(* CODESYS project listofinterface.library
   DefaultNamespace: KOSTAL.TC3.Components.ListOf.Interface
   DocFormat: reStructuredText
   Description: List of Items from base Interface {KOSTAL_TC3_Core_System.I_Interface}
      In addition to the interface, each item contains the pointer to the previous item as well as the pointer to the next item in the list.
   Author: Frank Dümpelmann
   Title: KOSTAL.TC3.Components.ListOf.Interface
   Version: 2019.1.0.0
   Company: KOSTAL GmbH & Co.KG
   Placeholder: KOSTAL.TC3.Components.ListOf.Interface

Project tree, tasks and I/O mapping:
  libraries: KOSTAL.TC3.Core.functionResponse, 2019.0.3.0 (KOSTAL GmbH & Co.KG); KOSTAL.TC3.Core.Settings, 2019.0.1.0 (KOSTAL GmbH & Co.KG); KOSTAL.TC3.Core.System, 2019.0.0.0 (KOSTAL GmbH & Co.KG); Tc2_Standard, 3.3.3.0 (Beckhoff Automation GmbH)
  0_Core/
    BaseElement/
      data type P_List
      data type ST_List
    function block FB_Core [ST]: _addItem, _findItem, _findItemByIndex, _insertItem, _removeFromBegin, _removeFromEnd, _removeItem, _removeItemByIndex, _nextItem, _previousItem, _clearResult, _setResultFail, _setResultPass, _checkConsistency, _clear, _NumberOfMember, _RegKey, FB_exit, FB_init
    interface I_Core
    interface I_Core_Owner
  1_Base/
    function block FB_Base [ST]: _verifyMember, _FIFO_peek, _FIFO_pop, _FIFO_push, _addMember, _findMember, _findMemberByIndex, _insertMember, _removeFromBegin, _removeFromEnd, _removeMember, _removeMemberByIndex, _clear, FB_exit, FB_init
    interface I_Base
    interface I_Base_Owner
  Project Information/
    function F_GetCompany [ST]
    function F_GetTitle [ST]
    function F_GetVersion [ST]
  Version/
    global variables Global_Version
*)

// 0_Core/BaseElement/P_List
//Pointer to an element of List
TYPE P_List : POINTER TO ST_List; END_TYPE

// 0_Core/BaseElement/ST_List
{attribute 'enable_dynamic_creation'}
TYPE ST_List :
	STRUCT
			pNext	 		: P_List;				//Pointer to next Item
			iMember		: KOSTAL_TC3_Core_System.I_Interface;	//Interface of this item
			pPrevious : P_List;				//Pointer to previous item
	END_STRUCT
END_TYPE

// Version/Global_Version
{attribute 'TcGenerated'}
{attribute 'no-analysis'}
{attribute 'linkalways'}
// This function has been automatically generated from the project information.
VAR_GLOBAL CONSTANT
	{attribute 'const_non_replaced'}
	stLibVersion_KOSTAL_TC3_Components_ListOf_Interface : ST_LibVersion := (iMajor := 2019, iMinor := 1, iBuild := 0, iRevision := 0, nFlags := 1, sVersion := '2019.1.0.0');
END_VAR

// 0_Core/FB_Core
(*

| =========================================================================
| List of Items from base Interface {KOSTAL_TC3_Core_System.I_Interface} 
| =========================================================================

..code::

	//In addition to the interface, each item contains the pointer to the previous item 
	//as well as the pointer to the next item in the list.

	TYPE ST_List :
		STRUCT
				pNext			: P_List;
				iMember		: KOSTAL_TC3_Core_System.I_Interface;	
				pPrevious : P_List;
		END_STRUCT
	END_TYPE

============= ======================================= ======================
| The List is defined by (p)Begin and (p)End and also the count of Members 
----------------------------------------------------------------------------
============= ======================================= ======================
 **_pBegin**  >>>>>>>>>>>>>>>>>>>>>>>>>>>>>>>>>>>>>>  **_pEnd**                     
 **Item-1**	    Item-2   Item-3   Item-4  Item-5      **Item-n**                   
============= ======================================= ======================



| =========================================================================
| The Member is an Interface as payload and an access pointer to the        
| previous member and the next member                                      
| ---------------------------------------------------------------------------
| Previous Item ---<<<Pointer-Previous-[Item]-Pointer-Next>>>---NextItem---
| =========================================================================

*)
FUNCTION_BLOCK ABSTRACT FB_Core IMPLEMENTS I_Core, I_Core_Owner

VAR
	_pBegin	: P_List;	//origin of List
  _pEnd		: P_List;	//end of List
	_Count	: UDINT;	//number of registered Member
	
	_RegKeyValue	: UDINT:= UDINT#0;	//use to create an unique ID
	
END_VAR

(*
	add new item to end of list
*)
METHOD PROTECTED _addItem : BOOL

VAR_INPUT
	Item		: KOSTAL_TC3_Core_System.I_Interface;
	Result	: REFERENCE TO KOSTAL_TC3_Core_functionResponse.FB_functionResponse;
END_VAR

VAR
	_pNewItem	: P_List;
END_VAR
_clearResult(Result);

IF Item = 0 THEN _setResultFail(Result, 'Parameter Item is empty');	RETURN;	END_IF


//create a new Item
_pNewItem:= __NEW(ST_List);

//If creation failed 
IF _pNewItem = 0 THEN _setResultFail(Result, 'New Item cannot create');	RETURN;	END_IF

//If list is empty
IF THIS^._Count = 0 (*THIS^._pEnd = 0*) THEN THIS^._pBegin:= THIS^._pEnd:= _pNewItem; 
ELSE

	//set new item previous item to actual last item (THIS^._pEnd)
	_pNewItem^.pPrevious:= THIS^._pEnd;
	_pNewItem^.pPrevious^.pNext:= _pNewItem;
 
	THIS^._pEnd:= _pNewItem;
END_IF

THIS^._pEnd^.iMember:= Item;
THIS^._Count:= THIS^._Count + UDINT#1;

_setResultPass(Result, 'addItem successful');

_RegKeyValue:= _RegKeyValue + 1;

_addItem:= TRUE;
END_METHOD

(*
	Search for the element {Item} in the list and return {FoundItem} if it is found {_findItem = TRUE}
*)
METHOD PROTECTED _findItem : BOOL
VAR_INPUT
	Item			: KOSTAL_TC3_Core_System.I_Interface;
	FoundItem	: REFERENCE TO P_List;
	Result		: REFERENCE TO KOSTAL_TC3_Core_functionResponse.FB_functionResponse;
END_VAR

VAR
	_Item		: P_List;
END_VAR

_clearResult(Result);

IF Item = 0 										THEN _setResultFail(Result, 'Parameter Item is empty');	RETURN;	END_IF
IF NOT __ISVALIDREF(FoundItem)	THEN _setResultFail(Result, 'FoundItem has no valid reference');	RETURN;	END_IF


_Item := THIS^._pBegin;

WHILE _Item <> 0 DO

	IF _Item^.iMember = Item THEN

		FoundItem := _Item;

		_findItem:= TRUE;

		_setResultPass(Result, 'Item found');
		
		RETURN;   

	END_IF
	
	_Item := THIS^._nextItem(_Item, 0);

END_WHILE

//FoundItem:= _Item;

_setResultFail(Result, 'Item not found');

_findItem:= FALSE;
END_METHOD

(*
	Search for the element {Item} in the list and return {FoundItem} if it is found {_findItem = TRUE}
*)
METHOD PROTECTED _findItemByIndex : BOOL
VAR_INPUT
	Index			: UDINT;
	FoundItem	: REFERENCE TO P_List;
	Result		: REFERENCE TO KOSTAL_TC3_Core_functionResponse.FB_functionResponse;
END_VAR

VAR
	_Item		: P_List;
	_udi: UDINT;
END_VAR

_findItemByIndex:= FALSE;

_clearResult(Result);

IF _Count = 0										THEN _setResultFail(Result, 'List is empty');											RETURN;	END_IF
IF Index > (_Count - 1)					THEN _setResultFail(Result, 'Parameter Index is out of range');		RETURN;	END_IF
IF NOT __ISVALIDREF(FoundItem)	THEN _setResultFail(Result, 'FoundItem has no valid reference');	RETURN;	END_IF


_Item := THIS^._pBegin;

IF Index > 0 THEN
	FOR _udi:= 0 TO Index - 1 DO
			_Item := THIS^._nextItem(_Item, 0);
	END_FOR
END_IF

FoundItem:= _Item;

IF FoundItem = 0 THEN
	_setResultFail(Result, 'Item not found');
ELSE	
	_setResultPass(Result, 'Item found');
	_findItemByIndex:= TRUE;
END_IF
END_METHOD

METHOD PROTECTED _insertItem : BOOL
VAR_INPUT
	Index		: UDINT;	//Index a which shall inserted the {Item}
	Item		: KOSTAL_TC3_Core_System.I_Interface;
	Result	: REFERENCE TO KOSTAL_TC3_Core_functionResponse.FB_functionResponse;
END_VAR

VAR
	_pNewItem			: P_List;
	_pExitingItem	: P_List;
END_VAR

_clearResult(Result);

//Item is empty
IF Item = 0 THEN _setResultFail(Result, 'Parameter Item is empty');	RETURN;	END_IF

//if List is empty add item 
IF (Index = 0) AND (_Count = 0)	THEN _insertItem:= _addItem(Item, Result);	RETURN;	END_IF

//Index is in list not available 
IF Index > (_Count - 1) THEN _setResultFail(Result, 'Index is out of range');	RETURN;	END_IF

//if index is end of list then add item to end of list 
IF (Index = (_Count - 1)) THEN _insertItem:= _addItem(Item, Result);	RETURN;	END_IF

//try to find item where shall inserted
IF NOT _findItemByIndex(Index, _pExitingItem, Result) THEN RETURN;	END_IF
IF _pExitingItem = 0 THEN _setResultFail(Result, 'Item not available');	RETURN;	END_IF


//create a new Item
_pNewItem:= __NEW(ST_List);

//If creation failed 
IF _pNewItem = 0 THEN _setResultFail(Result, 'New Item cannot create');	RETURN;	END_IF

_pNewItem^.iMember:= Item;

_pNewItem^.pNext		:= _pExitingItem;							//set the next item from new item to existing founded item
_pNewItem^.pPrevious:= _pExitingItem^.pPrevious;	//set the previous from existing item to the previous of new item

//if a previous exist then
//set the next from previous from existing item to the previous of new item
IF _pNewItem^.pPrevious <> 0 THEN	_pNewItem^.pPrevious^.pNext:= _pNewItem;	END_IF

_pExitingItem^.pPrevious:= _pNewItem;							//set the previous from existing founded item to  new item

//if inserted at the begin of list, set the begin pointer to new Item
IF THIS^._pBegin = _pExitingItem THEN	THIS^._pBegin:= _pNewItem;	END_IF

THIS^._Count:= THIS^._Count + UDINT#1;

_setResultPass(Result, 'insertItem successful');

_RegKeyValue:= _RegKeyValue + 1;

_insertItem:= TRUE;
END_METHOD

(*
	remove Item from begin of list
*)
METHOD PROTECTED _removeFromBegin : BOOL
VAR_INPUT
	Result	: REFERENCE TO KOSTAL_TC3_Core_functionResponse.FB_functionResponse;
END_VAR

_removeFromBegin:= THIS^._removeItemByIndex(0, Result);
END_METHOD

(*
	remove Item from end of list
*)
METHOD PROTECTED _removeFromEnd : BOOL
VAR_INPUT
	Result	: REFERENCE TO KOSTAL_TC3_Core_functionResponse.FB_functionResponse;
END_VAR

_removeFromEnd:= THIS^._removeItemByIndex(_Count, Result);
END_METHOD

(*
	remove given {Item} from List
*)
METHOD PROTECTED _removeItem : BOOL
VAR_INPUT
	Item		: P_List;
	Result	: REFERENCE TO KOSTAL_TC3_Core_functionResponse.FB_functionResponse;
END_VAR

_clearResult(Result);

IF Item = 0 THEN _setResultFail(Result, 'Parameter Item is empty');	RETURN;	END_IF

//exist a next member
IF Item^.pNext <> 0 THEN
	//set next members previous Item  to my previous Item
	Item^.pNext^.pPrevious := Item^.pPrevious; 
END_IF

//exist a previous member
IF Item^.pPrevious <> 0 THEN
	//set previous members next Item  to my next Item
	Item^.pPrevious^.pNext := Item^.pNext;
END_IF

//Item is the once member
IF Item = THIS^._pBegin AND Item = THIS^._pEnd THEN
	
	THIS^._pBegin := 0;
	THIS^._pEnd := 0;

ELSIF Item = THIS^._pBegin (*AND Item <> THIS^._pEnd*) THEN

	THIS^._pBegin := Item^.pNext;

ELSIF (*Item <> THIS^._pBegin AND*) Item = THIS^._pEnd THEN

	THIS^._pEnd := Item^.pPrevious;

END_IF

__DELETE(Item);

IF  THIS^._Count > UDINT#0 THEN	THIS^._Count := THIS^._Count - UDINT#1;	
ELSE
	_setResultFail(Result, 'removeItem Counter underflow');
	RETURN;
END_IF

_setResultPass(Result, 'removeItem successful');
_removeItem:= TRUE;
END_METHOD

(*
	remove given {Index} from List
*)
METHOD PROTECTED _removeItemByIndex : BOOL
VAR_INPUT
	Index		: UDINT;
	Result	: REFERENCE TO KOSTAL_TC3_Core_functionResponse.FB_functionResponse;
END_VAR

VAR
	_Item		: P_List;
	_bFound	: BOOL;
END_VAR

IF NOT _findItemByIndex(Index, _Item, Result)	THEN RETURN;	END_IF

_removeItemByIndex:= _removeItem(_Item, Result);
END_METHOD

// retreives the pointer to the next item of the given entry
METHOD PROTECTED _nextItem : P_List;
VAR_INPUT
    Item : P_List;
		Result	: REFERENCE TO KOSTAL_TC3_Core_functionResponse.FB_functionResponse;
END_VAR
VAR
	_Res	: P_List;
END_VAR

IF Item <> 0 THEN	_Res := Item^.pNext;
ELSE							_Res := 0;
END_IF

_nextItem:= _Res;
END_METHOD

// retreives the previous item of the given entry
METHOD PROTECTED _previousItem : P_List
VAR_INPUT
    Item 	: P_List;
END_VAR
VAR
	_Res	: P_List;
END_VAR

IF Item <> 0 THEN	_Res := Item^.pPrevious;
ELSE							_Res := 0;
END_IF

_previousItem:= _Res;
END_METHOD

(*
	Clear result component
*)
METHOD PROTECTED _clearResult : BOOL
VAR_INPUT
	IN : REFERENCE TO KOSTAL_TC3_Core_functionResponse.FB_functionResponse;
END_VAR

IF __ISVALIDREF(IN) THEN IN.clear(); _clearResult:= TRUE;	END_IF
END_METHOD

(*
	set result to fail with given information 
*)
METHOD PROTECTED _setResultFail : BOOL
VAR_INPUT
	IN : REFERENCE TO KOSTAL_TC3_Core_functionResponse.FB_functionResponse;
	Info	: KOSTAL_TC3_Core_Settings.T_MaxString;
END_VAR

IF __ISVALIDREF(IN) THEN 

	IN.success:= FALSE;
	IN.status:= Info;

	_setResultFail:= TRUE;

END_IF
END_METHOD

(*
	set result to pass with given information 
*)
METHOD PROTECTED _setResultPass : BOOL
VAR_INPUT
	IN : REFERENCE TO KOSTAL_TC3_Core_functionResponse.FB_functionResponse;
	Info	: KOSTAL_TC3_Core_Settings.T_MaxString;
END_VAR

IF __ISVALIDREF(IN) THEN 

	IN.success:= TRUE;
	IN.status:= Info;

	_setResultPass:= TRUE;

END_IF
END_METHOD

(*
	Check if the list is consistent
*)
METHOD PROTECTED _checkConsistency : BOOL
VAR_INPUT
	Result	: REFERENCE TO KOSTAL_TC3_Core_functionResponse.FB_functionResponse;
END_VAR

VAR
	_pItem			: P_List;
	_pNext			: P_List;
	_pPrev			: P_List;
	_nItemCounter	: UDINT;
	_bBeginOk			: BOOL;
	_bEndOk			: BOOL;
	_bPrevLinkOk		: BOOL;
	_bNextLinkOk		: BOOL;
	_bItemCountOk	: BOOL;
	_bInterfaceOk	: BOOL;
END_VAR
// check from pHead to pTail
_pItem:= THIS^._pBegin;
_nItemCounter:= 0;

IF THIS^._pBegin <> 0 THEN
	_bBeginOk:= (THIS^._pBegin^.pPrevious = 0);
ELSE
	_bBeginOk:= TRUE;
END_IF

IF THIS^._pEnd <> 0 THEN
	_bEndOk:= (THIS^._pEnd^.pNext = 0);
ELSE
	_bEndOk:= TRUE;
END_IF

IF _bBeginOk AND _bEndOk THEN

	_bPrevLinkOk:= TRUE;
	_bNextLinkOk:= TRUE;
	_bInterfaceOk:= TRUE;

	WHILE _pItem <> 0 DO
		
		_pPrev:= _pItem^.pPrevious;
		_pNext:= _pItem^.pNext;

		IF _pPrev <> 0 THEN
			_bPrevLinkOk:= (_pPrev^.pNext = _pItem);
		ELSE
			_bPrevLinkOk:= (_pItem = THIS^._pBegin);
		END_IF

		IF _pNext <> 0 THEN
			_bNextLinkOk:= (_pNext^.pPrevious = _pItem);
		ELSE
			_bNextLinkOk:= (_pItem = THIS^._pEnd);
		END_IF

		_bInterfaceOk:= (_pItem^.iMember <> 0);

		IF NOT _bNextLinkOk OR NOT _bPrevLinkOk OR NOT _bInterfaceOk THEN	EXIT;	END_IF

		//handle iteration
		_nItemCounter:= _nItemCounter + UDINT#1;
		_pItem:= THIS^._nextItem(_pItem, 0);

	END_WHILE

END_IF

_bItemCountOk:= (_nItemCounter = THIS^._Count);

IF 		NOT _bBeginOk			THEN	_setResultFail(Result, 'List head not ok');
ELSIF NOT _bEndOk				THEN	_setResultFail(Result, 'List End not ok');
ELSIF NOT _bPrevLinkOk 	THEN	_setResultFail(Result, Tc2_Standard.CONCAT('Previous Link failed by item ', UDINT_TO_STRING(_nItemCounter)));
ELSIF NOT _bNextLinkOk	THEN	_setResultFail(Result, Tc2_Standard.CONCAT('Next Link failed by item ', UDINT_TO_STRING(_nItemCounter)));
ELSIF NOT	_bInterfaceOk	THEN	_setResultFail(Result, Tc2_Standard.CONCAT('Interface failed by item ', UDINT_TO_STRING(_nItemCounter))); 
ELSIF NOT	_bItemCountOk THEN	_setResultFail(Result, 'Itemcounter is not ok');
ELSE													_setResultPass(Result, 'List is consistent');	_checkConsistency:= TRUE;
END_IF
END_METHOD

(*
	Delete the complete content of the list
*)
METHOD PROTECTED _clear

WHILE THIS^._pBegin <> 0 DO
    THIS^._removeItem(THIS^._pBegin, 0);  
END_WHILE
END_METHOD

//return the nnumber of items in List
PROPERTY PROTECTED _NumberOfMember : UDINT
GET

_NumberOfMember:= _Count;
END_GET
END_PROPERTY

PROPERTY PROTECTED _RegKey : UDINT
GET

_RegKey:= THIS^._RegKeyValue;
END_GET
END_PROPERTY

METHOD FB_exit : BOOL
VAR_INPUT
	bInCopyCode : BOOL; // if TRUE, the exit method is called for exiting an instance that is copied afterwards (online change).
END_VAR

_clear();
END_METHOD

METHOD FB_init : BOOL
VAR_INPUT
	bInitRetains : BOOL; // if TRUE, the retain variables are initialized (warm start / cold start)
	bInCopyCode : BOOL;  // if TRUE, the instance afterwards gets moved into the copy code (online change)
END_VAR

_clear();
END_METHOD

END_FUNCTION_BLOCK

// 0_Core/I_Core
INTERFACE I_Core EXTENDS KOSTAL_TC3_Core_System.I_Interface

END_INTERFACE

// 0_Core/I_Core_Owner
INTERFACE I_Core_Owner EXTENDS KOSTAL_TC3_Core_System.I_Interface

END_INTERFACE

// 1_Base/FB_Base
(*

| =========================================================================
| List of Items from base Interface {KOSTAL_TC3_Core_System.I_Interface} 
| =========================================================================

..code::

	//In addition to the interface, each item contains the pointer to the previous item 
	//as well as the pointer to the next item in the list.

	TYPE ST_List :
		STRUCT
				pNext			: P_List;
				iMember		: KOSTAL_TC3_Core_System.I_Interface;	
				pPrevious : P_List;
		END_STRUCT
	END_TYPE

============= ======================================= ======================
| The List is defined by (p)Begin and (p)End and also the count of Members 
----------------------------------------------------------------------------
============= ======================================= ======================
 **_pBegin**  >>>>>>>>>>>>>>>>>>>>>>>>>>>>>>>>>>>>>>  **_pEnd**                     
 **Item-1**	    Item-2   Item-3   Item-4  Item-5      **Item-n**                   
============= ======================================= ======================



| =========================================================================
| The Member is an Interface as payload and an access pointer to the        
| previous member and the next member                                      
| ---------------------------------------------------------------------------
| Previous Item ---<<<Pointer-Previous-[Item]-Pointer-Next>>>---NextItem---
| =========================================================================

*)
FUNCTION_BLOCK ABSTRACT FB_Base EXTENDS FB_Core IMPLEMENTS I_Base, I_Base_Owner

VAR
//	_pBegin	: P_List;	//origin of List
//  _pEnd		: P_List;	//end of List
//	_Count	: UDINT;	//number of registered Member
	
//	_RegKeyValue	: UDINT:= UDINT#0;	//use to create an unique ID
	
	//_Iterator 	: P_List;//???
END_VAR

(*
	integrate here the veryfing of your interface type 
	only if verifing is passed [_verifyMember:= TRUE] the called metode will proceeded 
*)
METHOD PROTECTED _verifyMember : BOOL

VAR_INPUT
	Member	: KOSTAL_TC3_Core_System.I_Interface;
	Result	: REFERENCE TO KOSTAL_TC3_Core_functionResponse.FB_functionResponse;
END_VAR

VAR
	_obj	: KOSTAL_TC3_Core_System.I_Interface;
	_bResult: BOOL;
END_VAR

IF Member = 0 THEN _setResultFail(Result, 'Parameter Member is empty');	RETURN;	END_IF

_bResult:= __QUERYINTERFACE(Member, _obj);

IF NOT _bResult OR (_obj = 0) THEN
	IF __ISVALIDREF(Result) THEN Result.success:= FALSE; Result.status:= 'no valid interface found';	END_IF	
	RETURN;
END_IF

_verifyMember:= TRUE;
END_METHOD

//methode return the Member from begin 
METHOD PROTECTED _FIFO_peek : BOOL
VAR_INPUT
	FoundMember	: REFERENCE TO KOSTAL_TC3_Core_System.I_Interface;	//return value
	Result			: REFERENCE TO KOSTAL_TC3_Core_functionResponse.FB_functionResponse;
END_VAR

_clearResult(Result);

IF 		NOT __ISVALIDREF(FoundMember) THEN _setResultFail(Result, 'FoundMember has no valid reference'); 
ELSE	_FIFO_peek:= _findMemberByIndex(0, FoundMember, Result);
END_IF
END_METHOD

//methode return the Member from begin and remove it from List
METHOD PROTECTED _FIFO_pop : BOOL
VAR_INPUT
	FoundMember	: REFERENCE TO KOSTAL_TC3_Core_System.I_Interface;	//return value
	Result			: REFERENCE TO KOSTAL_TC3_Core_functionResponse.FB_functionResponse;
END_VAR


_clearResult(Result);

_FIFO_pop:= _findMemberByIndex(0, FoundMember, Result);

IF _FIFO_pop THEN	_FIFO_pop:= _removeFromBegin(Result);	END_IF
END_METHOD

//push/add the {Member} to begin from List
METHOD PROTECTED _FIFO_push : BOOL
VAR_INPUT
	Member	: KOSTAL_TC3_Core_System.I_Interface;
	Result	: REFERENCE TO KOSTAL_TC3_Core_functionResponse.FB_functionResponse;
END_VAR


IF NOT _verifyMember(Member, Result)	THEN	RETURN;	END_IF

_FIFO_push:= _insertItem(UDINT#0, Member, Result);
END_METHOD

(*
	add new Member to end of list
*)
METHOD PROTECTED _addMember : BOOL

VAR_INPUT
	Member		: KOSTAL_TC3_Core_System.I_Interface;
	Result	: REFERENCE TO KOSTAL_TC3_Core_functionResponse.FB_functionResponse;
END_VAR


VAR
	_Member: KOSTAL_TC3_Core_System.I_Interface;
END_VAR

IF NOT _verifyMember(Member, Result)	THEN	RETURN;	END_IF

//member already exist
IF _findMember(Member,_Member, Result) THEN 
	_setResultFail(Result, 'The participant already exists in the list.');
	RETURN;	
END_IF	

_addMember:= _addItem(Member, Result);
END_METHOD

(*
	Search for the element {Item} in the list and return {FoundItem} if it is found {_findItem = TRUE}
*)
METHOD PROTECTED _findMember : BOOL
VAR_INPUT
	Member			: KOSTAL_TC3_Core_System.I_Interface;
	FoundMember	: REFERENCE TO KOSTAL_TC3_Core_System.I_Interface;	//return value
	Result			: REFERENCE TO KOSTAL_TC3_Core_functionResponse.FB_functionResponse;
END_VAR

VAR
	_Item		: P_List;
END_VAR

_clearResult(Result);

IF Member = 0 												THEN _setResultFail(Result, 'Parameter Item is empty');	RETURN;	END_IF
IF NOT __ISVALIDREF(FoundMember)			THEN _setResultFail(Result, 'FoundItem has no valid reference');	RETURN;	END_IF
IF NOT _verifyMember(Member, Result)	THEN	RETURN;	END_IF

_findMember:= _findItem(Member, _Item, Result);

IF NOT _findMember		THEN	RETURN;	END_IF
IF _Item = 0 					THEN	RETURN;	END_IF
//IF _Item^.iMember = 0 THEN	RETURN;	END_IF
IF NOT _verifyMember(_Item^.iMember, Result)	THEN	RETURN;	END_IF

FoundMember:= _Item^.iMember;
END_METHOD

//find a modul by index  
METHOD PROTECTED _findMemberByIndex : BOOL
VAR_INPUT
	Index				: UDINT;	//index of item
	FoundMember	: REFERENCE TO KOSTAL_TC3_Core_System.I_Interface;	//return value
	Result			: REFERENCE TO KOSTAL_TC3_Core_functionResponse.FB_functionResponse;	//result information
END_VAR

VAR
	_FoundItem	: P_List;
END_VAR

IF NOT __ISVALIDREF(FoundMember)	THEN _setResultFail(Result, 'FoundMember has no valid reference');	RETURN;	END_IF

FoundMember:= 0;

_findMemberByIndex:= _findItemByIndex(Index,_FoundItem, Result);

IF NOT _findMemberByIndex THEN RETURN;	END_IF

IF NOT _verifyMember(_FoundItem^.iMember, Result) THEN RETURN;	END_IF

FoundMember:= _FoundItem^.iMember;

_findMemberByIndex:= TRUE;
END_METHOD

METHOD PROTECTED _insertMember : BOOL
VAR_INPUT
	Index		: UDINT;	//Index a which shall inserted the {Item}
	Member	: KOSTAL_TC3_Core_System.I_Interface;
	Result	: REFERENCE TO KOSTAL_TC3_Core_functionResponse.FB_functionResponse;
END_VAR

VAR
	_Member: KOSTAL_TC3_Core_System.I_Interface;
END_VAR

IF NOT _verifyMember(Member, Result)	THEN	RETURN;	END_IF

//member already exist
IF _findMember(Member,_Member, Result) THEN 
	_setResultFail(Result, 'The participant already exists in the list.');
	RETURN;	
END_IF	

_insertMember:= _insertItem(Index, Member, Result);
END_METHOD

(*
	remove Item from begin of list
*)
METHOD PROTECTED _removeFromBegin : BOOL
VAR_INPUT
	Result	: REFERENCE TO KOSTAL_TC3_Core_functionResponse.FB_functionResponse;
END_VAR

_removeFromBegin:= THIS^._removeMemberByIndex(0, Result);
END_METHOD

(*
	remove Item from end of list
*)
METHOD PROTECTED _removeFromEnd : BOOL
VAR_INPUT
	Result	: REFERENCE TO KOSTAL_TC3_Core_functionResponse.FB_functionResponse;
END_VAR

_removeFromEnd:= THIS^._removeMemberByIndex(_Count, Result);
END_METHOD

(*
	remove given {Member} from List
*)
METHOD PROTECTED _removeMember : BOOL
VAR_INPUT
	Member	: KOSTAL_TC3_Core_System.I_Interface;
	Result	: REFERENCE TO KOSTAL_TC3_Core_functionResponse.FB_functionResponse;
END_VAR

VAR
	_Item		: P_List;
	_bFound: BOOL;
END_VAR


IF NOT _verifyMember(Member, Result)	THEN	RETURN;	END_IF

_bFound:= _findItem(Member, _Item, Result);

IF NOT _bFound THEN RETURN;	END_IF

_removeMember:= _removeItem(_Item, Result);
END_METHOD

(*
	remove given {Index} from List
*)
METHOD PROTECTED _removeMemberByIndex : BOOL
VAR_INPUT
	Index		: UDINT;
	Result	: REFERENCE TO KOSTAL_TC3_Core_functionResponse.FB_functionResponse;
END_VAR

VAR
	_bFound	: BOOL;
	_Member	: KOSTAL_TC3_Core_System.I_Interface;

END_VAR

IF NOT _findMemberByIndex(Index, _Member, Result)	THEN RETURN;	END_IF

_removeMemberByIndex:= _removeMember(_Member, Result);
END_METHOD

(*
	Delete the complete content of the list
*)
METHOD PROTECTED _clear
VAR_INPUT
END_VAR

WHILE THIS^._pBegin <> 0 DO
    THIS^._removeMember(THIS^._pBegin^.iMember, 0);  
END_WHILE
END_METHOD

METHOD FB_exit : BOOL
VAR_INPUT
	bInCopyCode : BOOL; // if TRUE, the exit method is called for exiting an instance that is copied afterwards (online change).
END_VAR

_clear();
END_METHOD

METHOD FB_init : BOOL
VAR_INPUT
	bInitRetains : BOOL; // if TRUE, the retain variables are initialized (warm start / cold start)
	bInCopyCode : BOOL;  // if TRUE, the instance afterwards gets moved into the copy code (online change)
END_VAR

_clear();
END_METHOD

END_FUNCTION_BLOCK

// 1_Base/I_Base
INTERFACE I_Base EXTENDS I_Core

END_INTERFACE

// 1_Base/I_Base_Owner
INTERFACE I_Base_Owner EXTENDS I_Core_Owner

END_INTERFACE

// Project Information/F_GetCompany
// This function has been automatically generated from the project information.
{attribute 'signature_flag' := '1073741824'}
{attribute 'TcGenerated'}
{attribute 'no-analysis'}
FUNCTION F_GetCompany : WSTRING
VAR_INPUT
	
END_VAR

F_GetCompany := "KOSTAL GmbH & Co.KG";

END_FUNCTION

// Project Information/F_GetTitle
// This function has been automatically generated from the project information.
{attribute 'signature_flag' := '1073741824'}
{attribute 'TcGenerated'}
{attribute 'no-analysis'}
FUNCTION F_GetTitle : WSTRING
VAR_INPUT
	
END_VAR

F_GetTitle := "KOSTAL.TC3.Components.ListOf.Interface";

END_FUNCTION

// Project Information/F_GetVersion
// This function has been automatically generated from the project information.
{attribute 'signature_flag' := '1073741824'}
{attribute 'TcGenerated'}
{attribute 'no-analysis'}
FUNCTION F_GetVersion : ST_LibVersion
VAR_INPUT
	
END_VAR

F_GetVersion.iMajor := 2019;
F_GetVersion.iMinor := 1;
F_GetVersion.iBuild := 0;
F_GetVersion.iRevision := 0;
F_GetVersion.sVersion := '2019.1.0.0';
F_GetVersion.nFlags := 1;

END_FUNCTION
